(* IEC 61131-3 sources: Lasal-MCP/examples/SampleSource/4_PumpControlSchemeSolution/Stations/MachineControl/MachineControl/Class/_SyncTimePLC, 1 file *)

(* ---- _SyncTimePLC.st ---- *)
#define SyncTimeDate 60sec

(*!
<Class
	Name               = "_SyncTimePLC"
	Revision           = "1.3"
	RealtimeTask       = "false"
	CyclicTask         = "false"
	DefCyclictime      = "60000 ms"
	BackgroundTask     = "true"
	DefBackground      = "30000 ms"
	Sigmatek           = "true"
	OSInterface        = "false"
	HighPriority       = "false"
	Automatic          = "false"
	UpdateMode         = "Prescan"
	SharedCommandTable = "true"
	Objectsize         = "(510,360)"
	Comment            = "sets every minute the source date &amp; time to the destination date &amp; time.&#13;&#10;(the values will be fixed by the background time)">
	<Channels>
		<Server Name="ClassSvr" Visualized="false" Initialize="false" WriteProtected="true" Retentive="false" Comment="class server"/>
		<Client Name="cOnline" Required="true" Internal="false" Comment="data channel to _MMStateSvr for reading the multimaster online status"/>
		<Client Name="cSetDate" Required="true" Internal="false" Comment="destination date"/>
		<Client Name="cSetTime" Required="true" Internal="false" Comment="destination time"/>
		<Client Name="cSyncDate" Required="true" Internal="false" Comment="source date "/>
		<Client Name="cSyncTime" Required="true" Internal="false" Comment="source time"/>
	</Channels>
	<Dependencies>
		<Files>
			<File Path=".\Class\_SyncTimePLC\_SyncTimePLC_en.pdf"/>
			<File Path=".\Class\_SyncTimePLC\_SyncTimePLC_de.pdf"/>
		</Files>
	</Dependencies>
	<RevDoku>
		<Owner Company="Sigmatek"/>
		<Dokumentation Revision="1.3" Date="2016-11-10" Author="KaiAnd" Company="Sigmatek" Description="changed type of client &quot;cOnline&quot; from &quot;_MMState&quot; to &quot;_SIG_LSL_CMultimasterState::_MMStateSvr&quot;&#13;&#10;(necessary because of changed type after action &quot;PROJECT -&gt; Multimaster -&gt; Create/Update State Class&quot;) "/>
		<Dokumentation Revision="1.2" Date="2016-10-10" Author="HubChr" Company="Sigmatek" Description="Added documentation pdfs."/>
		<Dokumentation Revision="1.1" Date="2016-09-07" Author="HubChr" Company="Sigmatek" Description="Translated comments to english"/>
		<Dokumentation Revision="1.0" Date="2015-11-11" Author="hötant" Company="Sigmatek" Description="creation of class"/>
	</RevDoku>
</Class>
*)
_SyncTimePLC : CLASS
  //Servers:
	ClassSvr 	: SvrChCmd_DINT;
  //Clients:
	cOnline 	: CltCh__MMStateSvr_PTofCls__SIG_LSL_CMultimasterState;
	cSyncDate 	: CltCh_HDINT;
	cSyncTime 	: CltCh_HDINT;
	cSetDate 	: CltCh_HDINT;
	cSetTime 	: CltCh_HDINT;
  //Variables:
		TimeStamp 	: UDINT;
  //Functions:

	FUNCTION VIRTUAL GLOBAL Background
		VAR_INPUT
			EAX 	: UDINT;
		END_VAR
		VAR_OUTPUT
			state (EAX) 	: UDINT;
		END_VAR;
  //Tables:
	FUNCTION @STD
		VAR_OUTPUT
			ret_code	: CONFSTATES;
		END_VAR;
	FUNCTION GLOBAL TAB @CT_;
END_CLASS;

FUNCTION VIRTUAL GLOBAL _SyncTimePLC::Background
	VAR_INPUT
		EAX 	: UDINT;
	END_VAR
	VAR_OUTPUT
		state (EAX) 	: UDINT;
	END_VAR

  cOnline := cOnline.Read();
  if (cOnline = _SIG_LSL_CMultimasterState::_MMStateSvr::Online) then
    case ClassSvr of
    0 : // Read Time from HMI
        cSyncTime := cSyncTime.Read();
        // Set Time of HMI to PLC
        cSetTime := cSyncTime ;
        cSetTime.Write (cSetTime);
        ClassSvr +=1;
        TimeStamp := ops.tAbsolute;

    1 : if ((ops.tAbsolute - TimeStamp ) >= 1sec) then
          // Read Date from HMI
          cSyncDate := cSyncDate.Read();
          // Set Date of HMI to PLC
          cSetDate := cSyncDate ;
          cSetDate.Write (cSetDate);
          ClassSvr +=1;
          TimeStamp := ops.tAbsolute;
        end_if;

    2 : // Update time cyclically
        if ((ops.tAbsolute - TimeStamp) >= (SyncTimeDate/2)) then
          // Read Time from HMI
          cSyncTime := cSyncTime.Read();
          // Set Time of HMI to PLC
          cSetTime := cSyncTime ;
          cSetTime.Write (cSetTime);
          ClassSvr +=1;
          TimeStamp := ops.tAbsolute;
        end_if;

    3 : // Update date cyclically
        if ((ops.tAbsolute - TimeStamp) >= (SyncTimeDate/2)) then
          // Read Date from HMI
          cSyncDate := cSyncDate.Read();
          // Set Date of HMI to PLC
          cSetDate := cSyncDate ;
          cSetDate.Write (cSetDate);
          ClassSvr :=2;
          TimeStamp := ops.tAbsolute;
        end_if;

    end_case;
  else
    ClassSvr :=0;
  end_if;

	state := READY;

END_FUNCTION
